Fanuc KAREL source: KO00041.KL

PROGRAM KO00041
%NOLOCKGROUP
%ENVIRONMENT MIR
VAR
  P1: POSITION
  P2: XYZWPREXT
  F: BOOLEAN
  OUT: POSITION
BEGIN
  F = TRUE
  OUT = MIRROR(P1, P2, F)
END KO00041
